Fanuc TP program (LS listing): Featur.LS

/PROG  Featur
/ATTR
OWNER		= MNEDITOR;
COMMENT		= "RoboDK sequence";
PROG_SIZE	= 0;
CREATE		= DATE 31-12-14  TIME 12:00:00;
MODIFIED	= DATE 31-12-14  TIME 12:00:00;
FILE_NAME	= Featur;
VERSION		= 0;
LINE_COUNT	= 32;
MEMORY_SIZE	= 0;
PROTECT		= READ_WRITE;
TCD:  STACK_SIZE	= 0,
      TASK_PRIORITY	= 50,
      TIME_SLICE	= 0,
      BUSY_LAMP_OFF	= 0,
      ABORT_REQUEST	= 0,
      PAUSE_REQUEST	= 0;
DEFAULT_GROUP	= 1,*,*,*,*;
CONTROL_CODE	= 00000000 00000000;
/MN
   1:  ! Program generated by VerticalBot Studio for Fanuc LR Mate 200 ;
   2:  ! iD on 25/10/2026 12:00:00 ;
   3:  ! Using nominal kinematics. ;
   4:  UFRAME_NUM=2 ;
   5:  ! UF2:100.0,-50.0,20.0,0.0,0.0,30.0 ;
   6:  UTOOL_NUM=1 ;
   7:  ! UT1:10.0,0.0,120.0,0.0,15.0,0.0 ;
   8:J P[1] 45% CNT5 ACC100 ;
   9:L P[2] 300mm/sec CNT5 ACC100 ;
  10:C P[3]
       P[4] 300mm/sec CNT5 ;
  11:L P[5] 50mm/sec CNT0 ACC100 ;
  12:L P[6] 300mm/sec FINE ACC100 ;
  13:  DO[3]=ON ;
  14:  DO_GRIP=OFF ;
  15:  WAIT DI[5]=ON ;
  16:  $WAITTMOUT=2000 ;
  17:  WAIT DI_PART=ON TIMEOUT, LBL[1] ;
  18:  MESSAGE[Timed out for LBL 1] ;
  19:  PAUSE ;
  20:  LBL[1] ;
  21:  WAIT  0.50(sec) ;
  22:  ! a comment line ;
  23:  MESSAGE[Hello operator] ;
  24:  CALL MyFunc ;
  25:  CALL SetRPM(5000) ;
  26:  RAW_CODE_LINE;
  27:  CALL SubPick ;
  28:  UTOOL_NUM=1 ;
  29:  ! UT1:10.0,0.0,120.0,0.0,15.0,0.0 ;
  30:  ! Attach to Tool 1 ;
  31:J P[7] 22% FINE ACC100 ;
  32:  PAUSE ;
/POS
P[1]{
   GP1:
    UF : 2, UT : 1,
	J1=    -20.000 deg,	J2=    10.000 deg,	J3=    -20.000 deg,
	J4=    30.000 deg,	J5=    -40.000 deg,	J6=    50.000 deg
};
P[2]{
   GP1:
    UF : 2, UT : 1,        CONFIG : 'F U T, 0, 0, 0',
	X =   332.153  mm,	Y =  -359.974  mm,	Z =   826.762  mm,
	W =   -51.647 deg,	P =     9.441 deg,	R =  -168.258 deg
};
P[3]{
   GP1:
    UF : 2, UT : 1,        CONFIG : 'F U T, 0, 0, 0',
	X =   286.258  mm,	Y =  -372.547  mm,	Z =   823.386  mm,
	W =   -52.463 deg,	P =     8.848 deg,	R =  -172.388 deg
};
P[4]{
   GP1:
    UF : 2, UT : 1,        CONFIG : 'F U T, 0, 0, 0',
	X =   205.710  mm,	Y =  -434.222  mm,	Z =   836.210  mm,
	W =   -50.828 deg,	P =    10.031 deg,	R =   177.880 deg
};
P[5]{
   GP1:
    UF : 2, UT : 1,        CONFIG : 'F U T, 0, 0, 0',
	X =   332.153  mm,	Y =  -359.974  mm,	Z =   826.762  mm,
	W =   -51.647 deg,	P =     9.441 deg,	R =  -168.258 deg
};
P[6]{
   GP1:
    UF : 2, UT : 1,        CONFIG : 'F U T, 0, 0, 0',
	X =   286.258  mm,	Y =  -372.547  mm,	Z =   823.386  mm,
	W =   -52.463 deg,	P =     8.848 deg,	R =  -172.388 deg
};
P[7]{
   GP1:
    UF : 2, UT : 1,
	J1=    -20.000 deg,	J2=    10.000 deg,	J3=    -20.000 deg,
	J4=    30.000 deg,	J5=    -40.000 deg,	J6=    50.000 deg
};
/END
